// TIA Portal V20 export
Screen "14_Alarm"  1319x30
  ScreenItem "ctlAlarmView" at 0,0 size 1319x30  Type=HmiAlarmControl
  ScreenItem "btnAlarmScreen" at 0,0 size 1319x30  Type=HmiButton
